ABB RAPID module: prc_project.modx

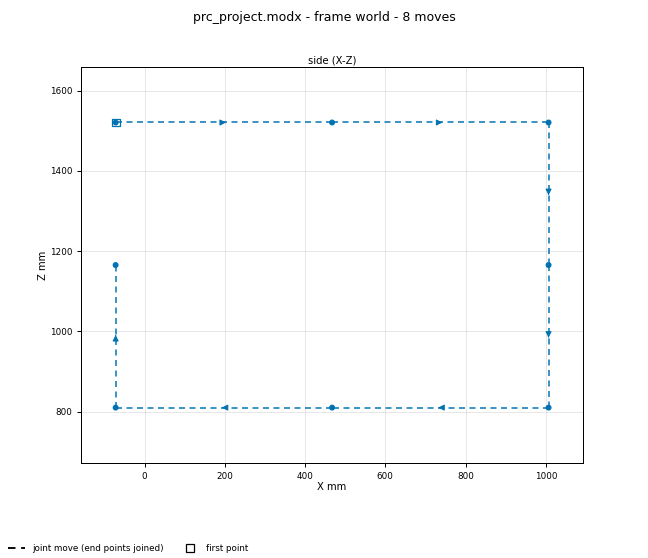
[picture p0: tool path of prc_project.modx in frame world, 8 of 10 moves have a stored position in this frame; points joined in program order, loops and branches not executed]
MODULE prc_project

    PERS wobjdata wobjBase := [
        FALSE, TRUE, "",
        [[0,0,0],[1,0,0,0]],
        [[0,0,0],[1,0,0,0]]
    ];
    PERS tooldata tool_0 := [
        TRUE,
        [[0,0,0],[1,0,0,0]],
        [0.001, [0,0,0.001], [1,0,0,0],0,0,0]
        ];

    PROC main()
        ConfL \Off;
        ConfJ \On;
        MoveAbsJ [[-90.000,0.000,20.000,0.000,-20.000,0.000], [9e9,9e9,9e9,9e9,9e9,9e9]], v500, fine, tool_0\WObj:=wobjBase;
        MoveJ [[-72.032,-2257.726,1520.434], [0.707107,0.707107,0.000000,0.000000], [-2,1,-1,0], [9e9,9e9,9e9,9e9,9e9,9e9]], v500, z50, tool_0\WObj:=wobjBase;
        MoveJ [[467.404,-2257.726,1520.434], [0.707107,0.707107,0.000000,0.000000], [-1,2,-2,0], [9e9,9e9,9e9,9e9,9e9,9e9]], v500, z50, tool_0\WObj:=wobjBase;
        MoveJ [[1006.839,-2257.726,1520.434], [0.707107,0.707107,0.000000,0.000000], [-1,2,-2,0], [9e9,9e9,9e9,9e9,9e9,9e9]], v500, z50, tool_0\WObj:=wobjBase;
        MoveJ [[1006.839,-2257.726,1165.192], [0.707107,0.707107,0.000000,0.000000], [-1,2,-2,0], [9e9,9e9,9e9,9e9,9e9,9e9]], v500, z50, tool_0\WObj:=wobjBase;
        MoveJ [[1006.839,-2257.726,809.950], [0.707107,0.707107,0.000000,0.000000], [-1,2,-2,0], [9e9,9e9,9e9,9e9,9e9,9e9]], v500, z50, tool_0\WObj:=wobjBase;
        MoveJ [[467.404,-2257.726,809.950], [0.707107,0.707107,0.000000,0.000000], [-1,2,-2,0], [9e9,9e9,9e9,9e9,9e9,9e9]], v500, z50, tool_0\WObj:=wobjBase;
        MoveJ [[-72.032,-2257.726,809.950], [0.707107,0.707107,0.000000,0.000000], [-2,1,-1,0], [9e9,9e9,9e9,9e9,9e9,9e9]], v500, z50, tool_0\WObj:=wobjBase;
        MoveJ [[-72.032,-2257.726,1165.192], [0.707107,0.707107,0.000000,0.000000], [-2,1,-1,0], [9e9,9e9,9e9,9e9,9e9,9e9]], v500, z50, tool_0\WObj:=wobjBase;
        MoveAbsJ [[-90.000,0.000,20.000,0.000,-20.000,0.000], [9e9,9e9,9e9,9e9,9e9,9e9]], v500, fine, tool_0\WObj:=wobjBase;
    ENDPROC
ENDMODULE
